{attribute 'no_assign'}
FUNCTION_BLOCK FB_LN_WTURBINE_LD0_WROT1 EXTENDS FB_AcsiCommonLogicalNodeClass
VAR_INPUT
	Beh: FB_DO_WTURBINE_LD0_WROT1_Beh := (sClass:='ENS', bLinkResult:=THIS^.AddDataToContainer(ipData:=Beh));
	RotSpd: FB_DO_WTURBINE_LD0_WROT1_RotSpd := (sClass:='MV', bLinkResult:=THIS^.AddDataToContainer(ipData:=RotSpd));
	BlPthAngTgt: FB_DO_WTURBINE_LD0_WROT1_BlPthAngTgt := (sClass:='MV', bLinkResult:=THIS^.AddDataToContainer(ipData:=BlPthAngTgt));
	BlPthAngVal: FB_DO_WTURBINE_LD0_WROT1_BlPthAngVal := (sClass:='MV', bLinkResult:=THIS^.AddDataToContainer(ipData:=BlPthAngVal));
END_VAR
VAR
END_VAR

END_FUNCTION_BLOCK

(* stored: Version 1.1.0.1
   POU FB_LN_WTURBINE_LD0_WROT1: Id {2ebb8303-e005-4174-88eb-1840d3b49d12}, SpecialFunc None *)
